Fanuc KAREL source: KA00136.KL

PROGRAM KA00136
%NOLOCKGROUP
VAR
  SRC: ARRAY[2] OF SHORT
  DST: STRING[80]
BEGIN
  SRC[1] = 2
  DST = SRC[1]
END KA00136
